Fanuc KAREL source: kt00438.KL

-- PROVISIONAL review KL for V1013-1; original PC SHA256 4c9aa2594ab5b7f98e6f567ee48047d1e774e40bb5e61ed6d312ff97f5629136
-- Incomplete behavior may be omitted. Consult companion uncertainty JSON. Do not deploy.
PROGRAM KT00438
%NOLOCKGROUP
VAR
  I1 : INTEGER
  R2 : REAL
  OUT : BOOLEAN
BEGIN
  -- UNRESOLVED_PC offsets 5-16; opcodes 2E,23
  -- UNRESOLVED_PC offsets 21-32; opcodes 2E,23
  -- UNRESOLVED_PC offsets 37-59; opcodes 21,21,29,64,29,72,23
  -- UNRESOLVED_PC offsets 64-68; opcodes 7F
END KT00438
